Fanuc KAREL source: kt00007.KL

-- PROVISIONAL review KL for V940-1; original PC SHA256 9f0082d9f9a6a578ec5ef99629727bccb1dfb04b09b6cb9b4e6371f0e3aaf40e
-- Incomplete behavior may be omitted. Consult companion uncertainty JSON. Do not deploy.
PROGRAM KT00007
%NOLOCKGROUP
VAR
  I1 : INTEGER
  OUT : INTEGER
-- UNRESOLVED_DECL H2 type=002017
BEGIN
  -- V9_ZERO_TABLE_METADATA_HINT layout=0001; no indexed target words; source/name/runtime held
  -- UNRESOLVED_PC offsets 5-16; opcodes 2E,23
  -- UNRESOLVED_PC offsets 21-35; opcodes 2E,22,9D,33,B4
  -- UNRESOLVED_PC offsets 40-62; opcodes 21,22,9D,33,B3,52,23
  -- UNRESOLVED_PC offsets 67-71; opcodes 7F
END KT00007
